Universal Robots URScript: T011_zai-org_GLM-4.7-FP8_baseline_rep2.urscript

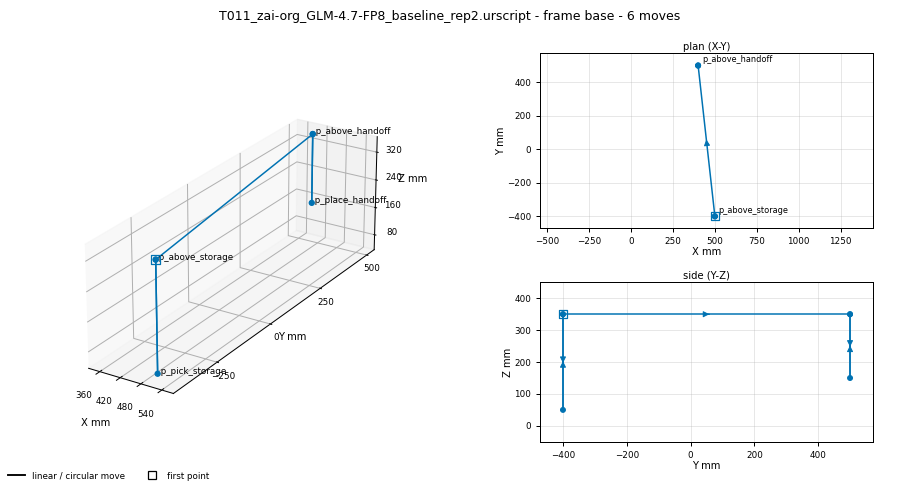
[picture p0: tool path of T011_zai-org_GLM-4.7-FP8_baseline_rep2.urscript in frame base, 6 of 8 moves have a stored position in this frame; points joined in program order, loops and branches not executed]
# Program: Dual-zone pick-place (T011)
# Robot: ur5e
# Mode: Hybrid
# Payload: 1.2 kg
# Description: Pick from fenced storage, place in collaborative handoff.

# Setup
set_payload(1.2, [0.0, 0.0, 0.05])
set_gravity([0.0, 0.0, 9.82])
set_tcp(p[0.0, 0.0, 0.0, 0.0, 0.0, 0.0])

# Define Poses
# Joint Home
q_home = [-1.57, -1.57, -1.57, -1.57, -1.57, 0.0]

# Storage Zone (Fenced - Industrial)
p_above_storage = p[0.5, -0.4, 0.35, 2.22, -2.22, 0.0]
p_pick_storage = p[0.5, -0.4, 0.05, 2.22, -2.22, 0.0]

# Handoff Zone (Collaborative - Operator)
p_above_handoff = p[0.4, 0.5, 0.35, 1.57, -3.14, 0.0]
p_place_handoff = p[0.4, 0.5, 0.15, 1.57, -3.14, 0.0]

# Move 1: move_joint: Home, 250.0 mm/s
movej(q_home, a=1.4, v=0.25, r=0)

# Move 2: move_linear: Above storage bin, 280.0 mm/s
movel(p_above_storage, a=1.2, v=0.28, r=0)

# Move 3: move_linear: Descend to pick, 120.0 mm/s
movel(p_pick_storage, a=0.5, v=0.12, r=0)

# gripper_action(pick)
set_digital_out(0, True)
sleep(0.5)

# Move 4: move_linear: Lift from bin, 200.0 mm/s
movel(p_above_storage, a=1.0, v=0.20, r=0)

# Move 5: move_linear: Transit to handoff zone, 250.0 mm/s
# Transitioning between zones (Hybrid mode logic applied via speed)
movel(p_above_handoff, a=1.2, v=0.25, r=0)

# Move 6: move_linear: Descend to handoff, 100.0 mm/s (Slower for safety)
movel(p_place_handoff, a=0.5, v=0.10, r=0)

# gripper_action(place)
set_digital_out(0, False)
sleep(0.5)

# Move 7: move_linear: Retract from handoff, 200.0 mm/s
movel(p_above_handoff, a=1.0, v=0.20, r=0)

# Move 8: move_joint: Return to Home, 250.0 mm/s
movej(q_home, a=1.4, v=0.25, r=0)

end
